Fanuc KAREL source: KT00712.KL

PROGRAM KT00712
%NOLOCKGROUP
VAR
  S1: STRING[80]
  S2: STRING[80]
  OUT: BOOLEAN
BEGIN
  S1 = 'A'
  S2 = 'B'
  S1 = 'A'
  S2 = 'B'
  OUT = UNINIT(S1)
END KT00712
